ABB RAPID module: TgtProg.mod

MODULE MainModule
GLOBAL VAR robtarget robpoint0= p:{{-607.850, 543.849, 363.215},{0.374108, 0.285846, 0.853660, -0.222712}}{cfg 0,0,0,4}{EJ 0.000000000,0.000000000,0.000000000,0.000000000,0.000000000,0.000000000}
GLOBAL VAR robtarget robpoint1= p:{{-607.850, 543.849, 363.215},{0.374108, 0.285846, 0.853660, -0.222712}}{cfg 0,0,0,2}{EJ 0.000000000,0.000000000,0.000000000,0.000000000,0.000000000,0.000000000}
GLOBAL VAR robtarget robpoint2= p:{{-607.850, 543.849, 363.215},{0.374108, 0.285846, 0.853660, -0.222712}}{cfg 0,0,0,7}{EJ 0.000000000,0.000000000,0.000000000,0.000000000,0.000000000,0.000000000}
GLOBAL VAR robtarget robpoint3= p:{{-607.850, 543.849, 363.215},{0.374108, 0.285846, 0.853660, -0.222712}}{cfg -1,-1,-1,0}{EJ 0.000000000,0.000000000,0.000000000,0.000000000,0.000000000,0.000000000}
GLOBAL VAR robtarget robpoint4= p:{{-607.850, 543.849, 363.215},{0.374108, 0.285846, 0.853660, -0.222712}}{cfg -2,3,2,0}{EJ 0.000000000,0.000000000,0.000000000,0.000000000,0.000000000,0.000000000}
GLOBAL VAR robtarget robpoint5= p:{{-607.850, 543.849, 363.215},{0.374108, 0.285846, 0.853660, -0.222712}}{cfg 2,4,-2,0}{EJ 0.000000000,0.000000000,0.000000000,0.000000000,0.000000000,0.000000000}

GLOBAL Proc main()
    MoveL robpoint0,v50,z50,tool03,wobj16
    MoveL robpoint1,v50,z50,tool03,wobj16
    MoveL robpoint2,v50,z50,tool03,wobj16
    MoveL robpoint3,v50,z50,tool03,wobj16
    MoveL robpoint4,v50,z50,tool03,wobj16
    MoveL robpoint5,v50,z50,tool03,wobj16
EndProc
EndModule
